// TIA Portal project "000_empty" (V21)

(* hardware
DEVICE "PLC_1"  S7-1500 station
   slot 0: "Rail_0"  Rack  6ES7 590-1***0-0AA0
   slot 1: "PLC_1"  CPU 1513-1 PN  6ES7 513-1AL02-0AB0  V2.9
      slot 3: "CPU display_1"  6ES7591-1AA00-0AA0
      slot 32768: "PROFINET interface_1"  X1
         slot 32769: "Port_1"  X1 P1
         slot 32770: "Port_2"  X1 P2
      slot 34817: "Virtual CP interface port_1"  Virtual CP interface port  Virtual CP interface port
*)

// ===== PLC "PLC_1"  CPU 1513-1 PN =====

TYPE "UDT_Motor"
   STRUCT
      Running : Bool;   // Motor on
      Speed : Real := 1500.0;   // Speed setpoint
      Count : Int := 7;
   END_STRUCT;
END_TYPE

DATA_BLOCK "DB_Global"   // DB1
{ S7_Optimized_Access := 'TRUE' }
   VAR
      xBool : Bool := TRUE;   // Bool comment
      iInt : Int := 42;
      rReal : Real := 3.5;   // Real comment
      aInt : Array[0..3] of Int;
      sData : Struct
         "a" : Bool;
         "b" : DInt := -5;
      END_STRUCT;
   END_VAR
BEGIN
   aInt[1] := 11;
END_DATA_BLOCK

DATA_BLOCK "FB_Empty_DB"   // DB2
{ S7_Optimized_Access := 'TRUE' }
VERSION : 0.1
// stored: InstanceOfName FB_Empty
"FB_Empty"
BEGIN
END_DATA_BLOCK

DATA_BLOCK "DB_Motor"   // DB4
{ S7_Optimized_Access := 'TRUE' }
   VAR
      motor : "UDT_Motor";
   END_VAR
BEGIN
   motor.Speed := 750.0;
END_DATA_BLOCK

DATA_BLOCK "FB_Iface_DB"   // DB5
{ S7_Optimized_Access := 'TRUE' }
VERSION : 0.1
// stored: InstanceOfName FB_Iface
"FB_Iface"
BEGIN
   stInt := 99;
   stBool := TRUE;
END_DATA_BLOCK

DATA_BLOCK "FB_SysMulti_DB"   // DB6
{ S7_Optimized_Access := 'TRUE' }
VERSION : 0.1
// stored: InstanceOfName FB_SysMulti
"FB_SysMulti"
BEGIN
END_DATA_BLOCK

DATA_BLOCK "DB_Buf"   // DB57
{ S7_Optimized_Access := 'TRUE' }
VERSION : 0.1
   VAR
      buf : Array[0..99] of Byte;
      "b" : Bool;
      w : Word;
      s : String;
   END_VAR
BEGIN
END_DATA_BLOCK

// folder: BlockGroup_1

DATA_BLOCK "DB_InGroup"   // DB3
{ S7_Optimized_Access := 'TRUE' }
   VAR
      wWord : Word := 16#00FF;
   END_VAR
BEGIN
END_DATA_BLOCK

// folder: System blocks/Program resources

DATA_BLOCK "DB_IEC_COUNTER"   // DB36
{ S7_Optimized_Access := 'TRUE' }
AUTHOR : Simatic
FAMILY : IEC
NAME : CNTR
VERSION : 1.0
// stored: InstanceOfName IEC_COUNTER
"IEC_COUNTER"
BEGIN
END_DATA_BLOCK

DATA_BLOCK "DB_IEC_DCOUNTER"   // DB37
{ S7_Optimized_Access := 'TRUE' }
AUTHOR : SIMATIC
FAMILY : IEC
NAME : DCNTR
VERSION : 1.2
// stored: InstanceOfName IEC_DCOUNTER
"IEC_DCOUNTER"
BEGIN
END_DATA_BLOCK

DATA_BLOCK "DB_IEC_LCOUNTER"   // DB38
{ S7_Optimized_Access := 'TRUE' }
AUTHOR : SIMATIC
FAMILY : IEC
NAME : LCNTR
VERSION : 1.2
// stored: InstanceOfName IEC_LCOUNTER
"IEC_LCOUNTER"
BEGIN
END_DATA_BLOCK

DATA_BLOCK "DB_IEC_LTIMER"   // DB39
{ S7_Optimized_Access := 'TRUE' }
AUTHOR : Simatic
FAMILY : IEC
NAME : IEC_LTMR
VERSION : 1.0
// stored: InstanceOfName IEC_LTIMER
"IEC_LTIMER"
BEGIN
END_DATA_BLOCK

DATA_BLOCK "DB_IEC_SCOUNTER"   // DB40
{ S7_Optimized_Access := 'TRUE' }
AUTHOR : Simatic
FAMILY : IEC
NAME : SCNTR
VERSION : 1.2
// stored: InstanceOfName IEC_SCOUNTER
"IEC_SCOUNTER"
BEGIN
END_DATA_BLOCK

DATA_BLOCK "DB_IEC_TIMER"   // DB41
{ S7_Optimized_Access := 'TRUE' }
AUTHOR : Simatic
FAMILY : IEC
NAME : IEC_TMR
VERSION : 1.0
// stored: InstanceOfName IEC_TIMER
"IEC_TIMER"
BEGIN
END_DATA_BLOCK

DATA_BLOCK "DB_IEC_UCOUNTER"   // DB42
{ S7_Optimized_Access := 'TRUE' }
AUTHOR : Simatic
FAMILY : IEC
NAME : UCNTR
VERSION : 1.2
// stored: InstanceOfName IEC_UCOUNTER
"IEC_UCOUNTER"
BEGIN
END_DATA_BLOCK

DATA_BLOCK "DB_IEC_UDCOUNTER"   // DB43
{ S7_Optimized_Access := 'TRUE' }
AUTHOR : Simatic
FAMILY : IEC
NAME : UDCNTR
VERSION : 1.2
// stored: InstanceOfName IEC_UDCOUNTER
"IEC_UDCOUNTER"
BEGIN
END_DATA_BLOCK

DATA_BLOCK "DB_IEC_ULCOUNTER"   // DB44
{ S7_Optimized_Access := 'TRUE' }
AUTHOR : Simatic
FAMILY : IEC
NAME : ULCNTR
VERSION : 1.2
// stored: InstanceOfName IEC_ULCOUNTER
"IEC_ULCOUNTER"
BEGIN
END_DATA_BLOCK

DATA_BLOCK "DB_IEC_USCOUNTER"   // DB45
{ S7_Optimized_Access := 'TRUE' }
AUTHOR : Simatic
FAMILY : IEC
NAME : USCNTR
VERSION : 1.2
// stored: InstanceOfName IEC_USCOUNTER
"IEC_USCOUNTER"
BEGIN
END_DATA_BLOCK

// folder: (top level)

FUNCTION_BLOCK "FB_Empty"   // FB1, SCL
{ S7_Optimized_Access := 'TRUE' }
VERSION : 0.1
BEGIN
END_FUNCTION_BLOCK

FUNCTION_BLOCK "FB_Iface"   // FB2, SCL
{ S7_Optimized_Access := 'TRUE' }
VERSION : 0.1
   VAR_INPUT
      iBool : Bool;   // Input bool
      iInt : Int;   // Input int
      iReal : Real;   // Input real
      iArr : Array[0..3] of Int;   // Input array
      iMotor : "UDT_Motor";   // Input UDT
   END_VAR
   VAR_OUTPUT
      oBool : Bool;   // Output bool
      oInt : Int;   // Output int
   END_VAR
   VAR_IN_OUT
      ioReal : Real;   // InOut real
   END_VAR
   VAR
      stInt : Int := 42;   // Static int
      stBool : Bool;   // Static bool comment
   END_VAR
   VAR_TEMP
      tInt : Int;   // Temp int
   END_VAR
   VAR CONSTANT
      cInt : Int := 7;   // Constant int
   END_VAR
BEGIN
   #tInt := #iInt + #cInt;
           #oInt := #tInt;
           #oBool := #iBool;
           #ioReal := #ioReal + #iReal;
END_FUNCTION_BLOCK

FUNCTION_BLOCK "FB_SysMulti"   // FB3, SCL
{ S7_Optimized_Access := 'TRUE' }
VERSION : 0.1
   VAR
      mTON_TIME : TON_TIME;
      mTOF_TIME : TOF_TIME;
      mTP_TIME : TP_TIME;
      mTONR_TIME : TONR_TIME;
      mTON_LTIME : TON_LTIME;
      mTOF_LTIME : TOF_LTIME;
      mTP_LTIME : TP_LTIME;
      mTONR_LTIME : TONR_LTIME;
      mCTU_INT : CTU_INT;
      mCTD_INT : CTD_INT;
      mCTUD_INT : CTUD_INT;
      mCTU_SINT : CTU_SINT;
      mCTU_DINT : CTU_DINT;
      mCTU_LINT : CTU_LINT;
      mCTU_UINT : CTU_UINT;
      mCTU_USINT : CTU_USINT;
      mCTU_UDINT : CTU_UDINT;
      mCTU_ULINT : CTU_ULINT;
      mCTD_DINT : CTD_DINT;
      mCTUD_DINT : CTUD_DINT;
      mCTUD_LINT : CTUD_LINT;
      mCTUD_UDINT : CTUD_UDINT;
      mR_TRIG : R_TRIG;
      mF_TRIG : F_TRIG;
      mTSEND_C : TSEND_C;
      mTRCV_C : TRCV_C;
      mTCON : TCON;
      mTDISCON : TDISCON;
      mTSEND : TSEND;
      mTRCV : TRCV;
      mTUSEND : TUSEND;
      mTURCV : TURCV;
      mTMAIL_C : TMAIL_C;
      mT_CONFIG : T_CONFIG;
      mGET : GET;
      mPUT : PUT;
      mUSEND : USEND;
      mURCV : URCV;
      mBSEND : BSEND;
      mBRCV : BRCV;
      mMB_CLIENT : MB_CLIENT;
      mMB_SERVER : MB_SERVER;
      mRDREC : RDREC;
      mWRREC : WRREC;
      mRALRM : RALRM;
      mGETIO : GETIO;
      mSETIO : SETIO;
      mGETIO_PART : GETIO_PART;
      mSETIO_PART : SETIO_PART;
      mProgram_Alarm : Program_Alarm;
      mDRUM : DRUM;
      mDCAT : DCAT;
      mMCAT : MCAT;
      mIMC : IMC;
      mSMC : SMC;
      mLEAD_LAG : LEAD_LAG;
      mPID_Compact : PID_Compact;
      mPID_3Step : PID_3Step;
      mPID_Temp : PID_Temp;
      mCONT_C : CONT_C;
      mCONT_S : CONT_S;
      mPULSEGEN : PULSEGEN;
      mTCONT_CP : TCONT_CP;
      mTCONT_S : TCONT_S;
      aTon : Array[0..1] of TON_TIME;
      aSend : Array[0..1] of TSEND_C;
   END_VAR
BEGIN
   #mTON_TIME(IN := TRUE, PT := T#1S);
END_FUNCTION_BLOCK

FUNCTION "FC_IecUse" : Void   // FC1, SCL
{ S7_Optimized_Access := 'TRUE' }
VERSION : 0.1
   VAR_INPUT
      "b" : Bool;
   END_VAR
BEGIN
   "DB_IEC_TIMER".TON(IN := #b, PT := T#1S);
   "DB_IEC_LTIMER".TON(IN := #b, PT := LT#1S);
   "DB_IEC_COUNTER".CTU(CU := #b, R := FALSE, PV := 5);
   "DB_IEC_SCOUNTER".CTU(CU := #b, R := FALSE, PV := 5);
   "DB_IEC_DCOUNTER".CTU(CU := #b, R := FALSE, PV := 5);
   "DB_IEC_LCOUNTER".CTU(CU := #b, R := FALSE, PV := 5);
   "DB_IEC_UCOUNTER".CTU(CU := #b, R := FALSE, PV := 5);
   "DB_IEC_USCOUNTER".CTU(CU := #b, R := FALSE, PV := 5);
   "DB_IEC_UDCOUNTER".CTU(CU := #b, R := FALSE, PV := 5);
   "DB_IEC_ULCOUNTER".CTU(CU := #b, R := FALSE, PV := 5);
END_FUNCTION

FUNCTION "FC_SysUse" : Void   // FC2, SCL
{ S7_Optimized_Access := 'TRUE' }
VERSION : 0.1
BEGIN
   "DB_TSEND_C"(CONNECT := "DB_Buf".buf, DATA := "DB_Buf".buf, ADDR := "DB_Buf".buf, COM_RST := "DB_Buf".b);
           "DB_TRCV_C"(CONNECT := "DB_Buf".buf, DATA := "DB_Buf".buf, ADDR := "DB_Buf".buf, COM_RST := "DB_Buf".b);
           "DB_TCON"(CONNECT := "DB_Buf".buf);
           "DB_TMAIL_C"(TO_S := "DB_Buf".s, CC := "DB_Buf".s, SUBJECT := "DB_Buf".s, TEXT := "DB_Buf".s, ATTACHMENT := "DB_Buf".buf, MAIL_ADDR_PARAM := "DB_Buf".buf);
           "DB_MB_CLIENT"(REQ := FALSE, DISCONNECT := FALSE, MB_MODE := 0, MB_DATA_ADDR := 0, MB_DATA_LEN := 0, MB_DATA_PTR := "DB_Buf".buf, CONNECT := "DB_Buf".buf, RD_MB_DATA_PTR := "DB_Buf".buf, WR_MB_DATA_PTR := "DB_Buf".buf);
           "DB_MB_SERVER"(MB_HOLD_REG := "DB_Buf".buf, CONNECT := "DB_Buf".buf);
           "DB_GETIO"(INPUTS := "DB_Buf".buf);
           "DB_SETIO"(OUTPUTS := "DB_Buf".buf);
           "DB_GETIO_PART"(INPUTS := "DB_Buf".buf);
           "DB_SETIO_PART"(OUTPUTS := "DB_Buf".buf);
           "DB_Program_Alarm"();
           "DB_DRUM"();
           "DB_DCAT"();
           "DB_MCAT"();
           "DB_IMC"();
           "DB_SMC"();
           "DB_LEAD_LAG"();
           "DB_PULSEGEN"();
           "DB_GET_SFB"(ADDR_1 := P#DB1.DBX0.0 BYTE 10, RD_1 := "DB_Buf".buf);
           "DB_PUT_SFB"(ADDR_1 := P#DB1.DBX0.0 BYTE 10, SD_1 := "DB_Buf".buf);
           "DB_RDREC_SFB"(RECORD := "DB_Buf".buf);
           "DB_WRREC_SFB"(RECORD := "DB_Buf".buf);
           "DB_RALRM_SFB"(TINFO := "DB_Buf".buf, AINFO := "DB_Buf".buf);
           "DB_T_CONFIG_SFB"();
           "DB_USEND_SFB"(SD_1 := "DB_Buf".buf, SD_2 := "DB_Buf".buf, SD_3 := "DB_Buf".buf, SD_4 := "DB_Buf".buf);
           "DB_URCV_SFB"(RD_1 := "DB_Buf".buf, RD_2 := "DB_Buf".buf, RD_3 := "DB_Buf".buf, RD_4 := "DB_Buf".buf);
           "DB_BSEND_SFB"(SD_1 := "DB_Buf".buf, LEN := "DB_Buf".w);
           "DB_BRCV_SFB"(RD_1 := "DB_Buf".buf, LEN := "DB_Buf".w);
           "DB_T_DISCON"();
           "DB_R_TRIG"();
           "DB_F_TRIG"();
END_FUNCTION

ORGANIZATION_BLOCK "Main"   // OB1, LAD, ProgramCycle
TITLE = "Main Program Sweep (Cycle)"
{ S7_Optimized_Access := 'TRUE' }
VERSION : 0.1
   VAR_INPUT
      Initial_Call : Bool;   // Initial call of this OB
      Remanence : Bool;   // =True, if remanent data are available
   END_VAR
BEGIN
END_ORGANIZATION_BLOCK